(* IEC 61131-3 sources: llm-plc-st-eval/data/processed_definitivo/gpt-4o-2024-08-06/C3/zero_shot, 3 files *)

(* ---- ejec_1.st ---- *)
PROGRAM PRG_Conversion
VAR
    // Declaración de variables de entrada
    btnMarcha : BOOL; // Botón de marcha
    btnParo : BOOL;   // Botón de paro

    // Declaración de variables de salida
    motor : BOOL;     // Estado del motor
    lampara : BOOL;   // Estado de la lámpara

    // Declaración del temporizador TON
    T1 : TON;         // Temporizador TON
END_VAR

// Lógica de control
// Rama 1: Control del motor
IF (btnMarcha OR motor) AND NOT btnParo THEN
    motor := TRUE;
ELSE
    motor := FALSE;
END_IF;

// Rama 2: Activación del temporizador TON
T1(IN := motor, PT := T#10S);

// Rama 3: Control de la lámpara
lampara := T1.Q;

(* ---- ejec_2.st ---- *)
PROGRAM PRG_Conversion
VAR
    btnMarcha : BOOL;   // Botón de marcha (entrada)
    btnParo : BOOL;     // Botón de paro (entrada)
    motor : BOOL;       // Estado del motor (salida)
    lampara : BOOL;     // Estado de la lámpara (salida)
    T1 : TON;           // Temporizador TON
END_VAR

// Lógica de control del motor
IF (btnMarcha OR motor) AND NOT btnParo THEN
    motor := TRUE;
ELSE
    motor := FALSE;
END_IF;

// Configuración y ejecución del temporizador TON
T1(IN := motor, PT := T#10S);

// Control de la lámpara basado en el temporizador
lampara := T1.Q;

(* ---- ejec_3.st ---- *)
PROGRAM PRG_Conversion
VAR
    // Entradas
    btnMarcha : BOOL; // Botón de marcha
    btnParo : BOOL;   // Botón de paro

    // Salidas
    motor : BOOL;     // Bobina del motor
    lampara : BOOL;   // Bobina de la lámpara

    // Temporizador
    T1 : TON;         // Temporizador TON
END_VAR

// Lógica de control
motor := (btnMarcha OR motor) AND NOT btnParo;

// Configuración y ejecución del temporizador
T1(IN := motor, PT := T#10S);

// Control de la lámpara
lampara := T1.Q;
